(* IEC 61131-3 sources: BioPrint-Automation-Suite/projects/02_bioprint_pid/plc/tests, 2 files *)

(* ---- FB_BioPrintPID_Test.st ---- *)
(* =============================================================================
   FB_BioPrintPID_Test — TcUnit test suite (TwinCAT 3; CODESYS via the TcUnit port)
   Replays the Python reference inputs scan by scan and checks every output.
   Instantiate in a PRG and call it cyclically, then call TcUnit.RUN().
   ============================================================================= *)
FUNCTION_BLOCK FB_BioPrintPID_Test EXTENDS TcUnit.FB_TestSuite
VAR
    fbPid       : FB_BioPrintPID;
    i           : INT;
    nMismatch   : INT;
    iFirst      : INT;
    lrWorst     : LREAL;
    lrDiff      : LREAL;
END_VAR

TEST('PID_ReplaysPythonReferenceVectors');

(* Start from a clean controller, defaults match config/default.toml *)
fbPid(bReset := TRUE);
fbPid.bReset := FALSE;

nMismatch := 0; iFirst := 0; lrWorst := 0.0;
FOR i := 1 TO GVL_ReferenceVectors.N_VECTORS DO
    fbPid(lrSetpoint    := GVL_ReferenceVectors.aPid[i].lrSetpoint,
          lrMeasurement := GVL_ReferenceVectors.aPid[i].lrMeasurement);
    lrDiff := ABS(fbPid.lrOutput - GVL_ReferenceVectors.aPid[i].lrOutput);
    lrWorst := MAX(lrWorst, lrDiff);
    IF lrDiff > 1.0E-6 THEN
        nMismatch := nMismatch + 1;
        IF iFirst = 0 THEN iFirst := i; END_IF;
    END_IF;
END_FOR;

AssertEquals_INT(Expected := 0, Actual := nMismatch,
    Message := CONCAT('output differs from Python by >1e-6 % duty; first scan ', INT_TO_STRING(iFirst)));
TEST_FINISHED();

TEST('PID_AntiWindupBoundsIntegrator');
fbPid(bReset := TRUE);
fbPid.bReset := FALSE;
FOR i := 1 TO 100 DO   (* 10 s pinned at 100 % with a 205 °C error *)
    fbPid(lrSetpoint := 230.0, lrMeasurement := 25.0);
END_FOR;
AssertTrue(Condition := fbPid.lrITerm <= 100.0, Message := 'integrator wound up past the output limit');
AssertTrue(Condition := fbPid.bSaturated, Message := 'saturation flag not set');
TEST_FINISHED();
END_FUNCTION_BLOCK

(* ---- FB_WestgardMonitor_Test.st ---- *)
(* =============================================================================
   FB_WestgardMonitor_Test — TcUnit test suite
   Replays the Python reference samples and checks every rule flag and the SD.
   ============================================================================= *)
FUNCTION_BLOCK FB_WestgardMonitor_Test EXTENDS TcUnit.FB_TestSuite
VAR
    fbQc      : FB_WestgardMonitor;
    i         : INT;
    nMismatch : INT;
    iFirst    : INT;
END_VAR

TEST('Westgard_ReplaysPythonReferenceVectors');

fbQc(bReset := TRUE, diStep := -1);
fbQc.bReset := FALSE;

nMismatch := 0; iFirst := 0;
FOR i := 1 TO GVL_ReferenceVectors.N_VECTORS DO
    fbQc(lrValue := GVL_ReferenceVectors.aWestgard[i].lrValue,
         diStep  := GVL_ReferenceVectors.aWestgard[i].diStep);
    IF fbQc.bWarn12s   <> GVL_ReferenceVectors.aWestgard[i].bWarn12s
    OR fbQc.bReject13s <> GVL_ReferenceVectors.aWestgard[i].bReject13s
    OR fbQc.bReject22s <> GVL_ReferenceVectors.aWestgard[i].bReject22s THEN
        nMismatch := nMismatch + 1;
        IF iFirst = 0 THEN iFirst := i; END_IF;
    END_IF;
END_FOR;

AssertEquals_LREAL(Expected := GVL_ReferenceVectors.LR_BASELINE_SD, Actual := fbQc.lrBaselineSd,
    Delta := 1.0E-9, Message := 'baseline SD differs from Python');
AssertEquals_INT(Expected := 0, Actual := nMismatch,
    Message := CONCAT('rule flags differ from Python; first sample ', INT_TO_STRING(iFirst)));
AssertTrue(Condition := fbQc.bRunRejected, Message := 'disturbance should reject the run');
TEST_FINISHED();
END_FUNCTION_BLOCK
